(* IEC 61131-3 sources: llm-plc-st-eval/data/processed_definitivo/claude-sonnet-4-6/I1/few_shot, 3 files *)

(* ---- ejec_1.st ---- *)
FUNCTION_BLOCK FB_Semaforo
VAR_INPUT
    habilitado : BOOL; (* Habilitacion del semaforo *)
END_VAR
VAR_OUTPUT
    luzV : BOOL; (* Luz verde *)
    luzA : BOOL; (* Luz amarilla *)
    luzR : BOOL; (* Luz roja *)
END_VAR
VAR
    estado      : INT;  (* Estado de la secuencia: 0=Verde, 1=Amarillo, 2=Rojo *)
    tFase       : TON;  (* Temporizador de fase normal *)
    tParpadeo   : TP;   (* Temporizador de pulso para amarillo intermitente *)
    bParpadeoOn : BOOL; (* Bandera de ciclo de parpadeo activo *)
END_VAR

IF NOT habilitado THEN
    (* --- Modo inhabilitado: amarillo intermitente 1s ON / 1s OFF --- *)
    estado := 0;        (* Reinicio de estado para cuando se habilite de nuevo *)
    tFase(IN := FALSE, PT := T#20S); (* Resetea temporizador de fase *)

    (* Genera el parpadeo usando TP: cada vez que Q baja, relanza el pulso *)
    tParpadeo(IN := NOT tParpadeo.Q AND NOT bParpadeoOn, PT := T#1S);

    (* Alterna entre encendido y apagado cada segundo *)
    IF tParpadeo.Q THEN
        bParpadeoOn := NOT bParpadeoOn;
    END_IF;

    luzV := FALSE;
    luzA := bParpadeoOn; (* Amarillo parpadea *)
    luzR := FALSE;

ELSE
    (* --- Modo habilitado: secuencia Verde -> Amarillo -> Rojo --- *)
    tParpadeo(IN := FALSE, PT := T#1S); (* Resetea temporizador de parpadeo *)
    bParpadeoOn := FALSE;

    CASE estado OF

        0: (* Verde durante 20 segundos *)
            luzV := TRUE;
            luzA := FALSE;
            luzR := FALSE;
            tFase(IN := TRUE, PT := T#20S);
            IF tFase.Q THEN
                tFase(IN := FALSE, PT := T#20S); (* Resetea temporizador *)
                estado := 1;
            END_IF;

        1: (* Amarillo durante 4 segundos *)
            luzV := FALSE;
            luzA := TRUE;
            luzR := FALSE;
            tFase(IN := TRUE, PT := T#4S);
            IF tFase.Q THEN
                tFase(IN := FALSE, PT := T#4S); (* Resetea temporizador *)
                estado := 2;
            END_IF;

        2: (* Rojo durante 15 segundos *)
            luzV := FALSE;
            luzA := FALSE;
            luzR := TRUE;
            tFase(IN := TRUE, PT := T#15S);
            IF tFase.Q THEN
                tFase(IN := FALSE, PT := T#15S); (* Resetea temporizador *)
                estado := 0; (* Reinicia la secuencia en verde *)
            END_IF;

        ELSE
            estado := 0; (* Estado invalido: vuelve a verde *)

    END_CASE;

END_IF;

END_FUNCTION_BLOCK

(* ---- ejec_2.st ---- *)
FUNCTION_BLOCK FB_Semaforo
VAR_INPUT
    habilitado : BOOL; (* Habilita la secuencia normal del semaforo *)
END_VAR
VAR_OUTPUT
    luzV : BOOL; (* Luz verde *)
    luzA : BOOL; (* Luz amarilla *)
    luzR : BOOL; (* Luz roja *)
END_VAR
VAR
    estado     : INT;  (* Estado de la secuencia: 0=Verde, 1=Amarillo, 2=Rojo *)
    tFase      : TON; (* Temporizador de cada fase de la secuencia normal *)
    tBlink     : TP;  (* Temporizador de pulso para amarillo intermitente *)
    blink      : BOOL; (* Estado actual del parpadeo amarillo *)
    prevHab    : BOOL; (* Valor anterior de habilitado para detectar flancos *)
END_VAR

IF habilitado THEN
    (* --- Secuencia normal: Verde -> Amarillo -> Rojo -> (repite) --- *)

    (* Al detectar flanco ascendente de habilitado, reiniciar en verde *)
    IF NOT prevHab THEN
        estado := 0;
        tFase(IN := FALSE, PT := T#20S); (* Reset del temporizador *)
    END_IF;

    CASE estado OF

        0: (* VERDE: 20 segundos *)
            tFase(IN := TRUE, PT := T#20S);
            luzV := TRUE;
            luzA := FALSE;
            luzR := FALSE;
            IF tFase.Q THEN
                tFase(IN := FALSE, PT := T#20S); (* Reset *)
                estado := 1;
            END_IF;

        1: (* AMARILLO: 4 segundos *)
            tFase(IN := TRUE, PT := T#4S);
            luzV := FALSE;
            luzA := TRUE;
            luzR := FALSE;
            IF tFase.Q THEN
                tFase(IN := FALSE, PT := T#4S); (* Reset *)
                estado := 2;
            END_IF;

        2: (* ROJO: 15 segundos *)
            tFase(IN := TRUE, PT := T#15S);
            luzV := FALSE;
            luzA := FALSE;
            luzR := TRUE;
            IF tFase.Q THEN
                tFase(IN := FALSE, PT := T#15S); (* Reset *)
                estado := 0; (* Reinicia ciclo en verde *)
            END_IF;

        ELSE
            estado := 0; (* Estado invalido: volver a verde *)

    END_CASE;

    (* Asegurar que el temporizador de parpadeo quede inactivo *)
    tBlink(IN := FALSE, PT := T#1S);
    blink := FALSE;

ELSE
    (* --- Modo inhabilitado: amarillo intermitente 1s ON / 1s OFF --- *)

    (* Apagar verde y rojo *)
    luzV := FALSE;
    luzR := FALSE;

    (* Asegurar que el temporizador de secuencia quede inactivo *)
    tFase(IN := FALSE, PT := T#20S);

    (* Generar pulso de 1 segundo repetitivo para el parpadeo *)
    tBlink(IN := NOT tBlink.Q, PT := T#1S);

    (* El pulso activo indica amarillo encendido *)
    luzA := tBlink.Q;

END_IF;

(* Guardar estado actual de habilitado para deteccion de flanco en proximo ciclo *)
prevHab := habilitado;

END_FUNCTION_BLOCK

(* ---- ejec_3.st ---- *)
FUNCTION_BLOCK FB_Semaforo
VAR_INPUT
    habilitado : BOOL; (* Habilita la secuencia normal del semaforo *)
END_VAR
VAR_OUTPUT
    luzV : BOOL; (* Luz verde *)
    luzA : BOOL; (* Luz amarilla *)
    luzR : BOOL; (* Luz roja *)
END_VAR
VAR
    estado     : INT;  (* Estado de la secuencia: 0=verde, 1=amarillo, 2=rojo *)
    tFase      : TON; (* Temporizador de cada fase normal *)
    tBlink     : TP;  (* Temporizador de pulso para amarillo intermitente *)
    bBlinkTrig : BOOL; (* Flanco para relanzar el pulso intermitente *)
END_VAR

IF habilitado THEN
    (* --- Secuencia normal: verde -> amarillo -> rojo -> verde --- *)

    CASE estado OF

        0: (* VERDE 20 s *)
            luzV := TRUE;
            luzA := FALSE;
            luzR := FALSE;
            tFase(IN := TRUE, PT := T#20S);
            IF tFase.Q THEN
                tFase(IN := FALSE, PT := T#20S); (* Resetea temporizador *)
                estado := 1;
            END_IF;

        1: (* AMARILLO 4 s *)
            luzV := FALSE;
            luzA := TRUE;
            luzR := FALSE;
            tFase(IN := TRUE, PT := T#4S);
            IF tFase.Q THEN
                tFase(IN := FALSE, PT := T#4S);
                estado := 2;
            END_IF;

        2: (* ROJO 15 s *)
            luzV := FALSE;
            luzA := FALSE;
            luzR := TRUE;
            tFase(IN := TRUE, PT := T#15S);
            IF tFase.Q THEN
                tFase(IN := FALSE, PT := T#15S);
                estado := 0; (* Reinicia ciclo *)
            END_IF;

        ELSE
            estado := 0; (* Estado invalido: vuelve a verde *)

    END_CASE;

    (* Asegura que el temporizador de blink quede inactivo *)
    bBlinkTrig := FALSE;
    tBlink(IN := FALSE, PT := T#1S);

ELSE
    (* --- Modo inhabilitado: amarillo intermitente 1 s ON / 1 s OFF --- *)
    luzV := FALSE;
    luzR := FALSE;

    (* Relanza el pulso cada vez que expira *)
    tBlink(IN := bBlinkTrig, PT := T#1S);

    IF NOT tBlink.Q AND NOT bBlinkTrig THEN
        (* Pulso inactivo y no disparado: lanzar nuevo pulso *)
        bBlinkTrig := TRUE;
    END_IF;

    IF tBlink.Q THEN
        (* Pulso expirado: apagar disparo para permitir nuevo ciclo *)
        bBlinkTrig := FALSE;
    END_IF;

    luzA := tBlink.Q; (* Amarillo encendido durante el pulso activo *)

    (* Al rehabilitar, reinicia la secuencia en verde *)
    tFase(IN := FALSE, PT := T#20S);
    estado := 0;

END_IF;

END_FUNCTION_BLOCK
